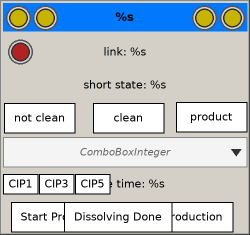
VISUALIZATION vis_FB_Element  // 250x235
VAR_IN_OUT
	fb: FB_Element;
END_VAR
    Rectangle (0,0 250x235)
    Textfield (3,70 244x30), "short state: %s", text variable: fb.eState_Short
    ComboBoxInteger (3,137 244x30), variable: fb.eState_Long, input disabled if: fb.bStateUpdate_Limited, text list: 'TextList_StateLong'
    Textfield (2,2 246x30), "%s", text variable: fb.sElementID
    Textfield (2,169 246x30), "state time: %s", text variable: fb.sState_Time
    RoundedRectangle (11,202 108x30), "Start Production", invisible if: NOT (fb.eInterConnect=E_InterConnection.ConnToLine AND fb.eState_Long=E_Element_State_Long.eReady)
        OnMouseClick: execute { fb.eState_Long:=E_Element_State_Long.eProduction; }
    RoundedRectangle (125,202 108x30), "Stop Production", invisible if: NOT (fb.eInterConnect=E_InterConnection.ConnToLine AND fb.eState_Long=E_Element_State_Long.eProduction)
        OnMouseClick: execute { fb.eState_Long:=E_Element_State_Long.eReady; }
    RoundedRectangle (64,202 108x30), "Dissolving Done", invisible if: NOT ((fb.eInterConnect=E_InterConnection.ConnToTriBlender) AND (fb.eState_Long=E_Element_State_Long.eCIP_5_Done OR fb.eState_Long=E_Element_State_Long.eWaterReady))
        OnMouseClick: execute { fb.eState_Long:=E_Element_State_Long.eReady; }
    Lamp1 (190,4 29x28), variable: fb.eInterConnect=E_InterConnection.ConnToLine, style: Lamp-Lamp1-Yellow
    Lamp1 (218,4 29x28), variable: fb.eInterConnect=E_InterConnection.ConnToTriBlender, style: Lamp-Lamp1-Yellow
    Lamp1 (31,4 29x28), variable: fb.eInterConnect=E_InterConnection.ConnToTank, style: Lamp-Lamp1-Yellow
    Textfield (3,37 244x30), "link: %s", colour toggle: fb.eInterConnect<>0, text list: 'TextList_InterConnection', text index: fb.eInterConnect
    RoundedRectangle (4,103 71x30), "not clean"
        OnMouseClick: execute { fb.eState_Long:=E_Element_State_Long.eNotClean; }
    RoundedRectangle (93,103 71x30), "clean"
        OnMouseClick: execute { fb.eState_Long:=E_Element_State_Long.eCIP_5_Done; }
    RoundedRectangle (176,102 71x30), "product"
        OnMouseClick: execute { fb.eState_Long:=E_Element_State_Long.eProduction; }
    Lamp1 (4,4 29x28), variable: fb.eInterConnect=E_InterConnection.ConnToCIP, style: Lamp-Lamp1-Yellow
    RoundedRectangle (3,174 35x20), "CIP1"
        tap fb.bTakePosInCIPBuffer_Partial
    RoundedRectangle (39,174 35x20), "CIP3"
        tap fb.bTakePosInCIPBuffer_Detergent
    RoundedRectangle (75,174 35x20), "CIP5"
        tap fb.bTakePosInCIPBuffer_Full
    Lamp1 (6,38 29x28), variable: fb.bError, style: Lamp-Lamp1-Red
END_VISUALIZATION

(* stored: Version 1.1.0.1, ProductVersion 3.1.4024.15
   Visu vis_FB_Element: Id {16669df6-d834-41fd-adf0-1a813ab2bb8a} *)
